{attribute 'qualified_only'}
TYPE E_AnalogOutputCommand : (NONE := 0, SET := 1) DINT;
END_TYPE

(* stored: Version 1.1.0.1, ProductVersion 3.1.4024.12
   DUT E_AnalogOutputCommand: Id {b4d42d0a-9eee-4c6f-acc2-7cc706f6f1fa} *)
